Staubli VAL3: main.pgx

program main()
begin
  close(tCurrentTool)
  pPointRs.config.shoulder = lefty
  pPointRs2.config.shoulder = lefty
  mCurrentSpeed.tvel = 100.00
  mCurrentSpeed.blend = joint
  mCurrentSpeed.reach = 0.010
  mCurrentSpeed.leave = 0.010
  // Program ManyMoves start
  // Program generated by RoboDK v6.0.7 for Staubli TP80 on XX/XX/XXXX 18:00:00
  // Using nominal kinematics.
  mCurrentSpeed.tvel = 500.000
  call MoveJoint(10.00000,-20.00000,50.00000,30.00000)
  call MoveLine(-638.084,504.480,372.034,136.262,30.757,-130.375)
  call MoveJoint(30.00000,25.00000,80.00000,-45.00000)
  // Linear movement using joint targets is not supported. Change the target type to cartesian or use a joint movement.
  call MoveJoint(10.00000,-20.00000,50.00000,30.00000)
  call MoveLine(-628.084,494.480,374.034,136.262,30.757,-130.375)
  call MoveJoint(30.00000,25.00000,80.00000,-45.00000)
  // Linear movement using joint targets is not supported. Change the target type to cartesian or use a joint movement.
  call MoveJoint(10.00000,-20.00000,50.00000,30.00000)
  call MoveLine(-618.084,484.480,376.034,136.262,30.757,-130.375)
  call MoveJoint(30.00000,25.00000,80.00000,-45.00000)
  // Linear movement using joint targets is not supported. Change the target type to cartesian or use a joint movement.
  call MoveJoint(10.00000,-20.00000,50.00000,30.00000)
  call MoveLine(-608.084,474.480,378.034,136.262,30.757,-130.375)
  call MoveJoint(30.00000,25.00000,80.00000,-45.00000)
  // Linear movement using joint targets is not supported. Change the target type to cartesian or use a joint movement.
  call MoveJoint(10.00000,-20.00000,50.00000,30.00000)
  call MoveLine(-598.084,464.480,380.034,136.262,30.757,-130.375)
  call MoveJoint(30.00000,25.00000,80.00000,-45.00000)
  // Linear movement using joint targets is not supported. Change the target type to cartesian or use a joint movement.
  call MoveJoint(10.00000,-20.00000,50.00000,30.00000)
  call MoveLine(-588.084,454.480,382.034,136.262,30.757,-130.375)
  call MoveJoint(30.00000,25.00000,80.00000,-45.00000)
  // Linear movement using joint targets is not supported. Change the target type to cartesian or use a joint movement.
  call MoveJoint(10.00000,-20.00000,50.00000,30.00000)
  call MoveLine(-578.084,444.480,384.034,136.262,30.757,-130.375)
  call MoveJoint(30.00000,25.00000,80.00000,-45.00000)
  // Linear movement using joint targets is not supported. Change the target type to cartesian or use a joint movement.
  call MoveJoint(10.00000,-20.00000,50.00000,30.00000)
  call MoveLine(-568.084,434.480,386.034,136.262,30.757,-130.375)
  call MoveJoint(30.00000,25.00000,80.00000,-45.00000)
  // Linear movement using joint targets is not supported. Change the target type to cartesian or use a joint movement.
  call MoveJoint(10.00000,-20.00000,50.00000,30.00000)
  call MoveLine(-558.084,424.480,388.034,136.262,30.757,-130.375)
  call MoveJoint(30.00000,25.00000,80.00000,-45.00000)
  // Linear movement using joint targets is not supported. Change the target type to cartesian or use a joint movement.
  call MoveJoint(10.00000,-20.00000,50.00000,30.00000)
  call MoveLine(-548.084,414.480,390.034,136.262,30.757,-130.375)
  call MoveJoint(30.00000,25.00000,80.00000,-45.00000)
  // Linear movement using joint targets is not supported. Change the target type to cartesian or use a joint movement.

  waitEndMove()
  // Program ManyMoves end

end
